LAYER ETE_TJ
  (* CLP SUBESTACAO (M262_Substacao) *)
  (* CLP LODO (M262_Lodo) *)
  (* CLP NEREDA (M262_Nereda) *)
  (* Painel Subestacao - Remota 1 (SUB_R1 .192), geradores QTAM1/QTAM2 (AGC150 .186/.187), MGE QGBT 220 V (.191) *)
  (* Agua de Reuso (1000) - Remota 2 (SUB_R2 .193), MGE .190 *)
  (* EEE Bruto (100) - Remota A1 (.197), inversores BS-100-01/02/03 (.200-.202), MGE .199 *)
  (* Pre-tratamento (200) - UCT_200_01 (.182), UCT_200_02 (.184), UCT_200_03 reserva; inversores BR-200-03/04 (.176/.177) *)
  (* Remota 2 do Nereda (NER_R2 .161, A12 canal 7) - lida pelo CLP Subestacao *)
  (* Gradeamento (100) - painel Vibropac (.207), comportas CO-100-01..04 (.203-.206) *)
  (* Sem painel definido - Dosagem de alcalinizante (800), sem campo *)
  (* Desinfeccao (700) - Remota A1, VC-700-01, UV Trojan, SC4500 pH/OD/turbidez, MGE .139 *)
  (* Lodo (900) - Remotas A2 (.135) e A10 (.136), inversores, valvulas e skids 900, MGE .246 *)
  (* Painel Nereda - Remotas A2/A10, Remota A11 (area do lodo: SludgeBuffer e Sludge Holding Tanks), sopradores Sulzer V4601-4604, SC1000/SC4500, inversores P4001-3/R4005/P4901-3, MGE .143 *)
  (* NEREDA REACTORS *)
  (* NEREDA PROCESS - HIDRYCO *)
  (* EMERGENCY RECIPIE *)
  (* NEREDA EQUIPMENT *)
  (* NEREDA AERATION *)
  (* INFLUENT FEED *)
  (* EFFLUENT *)
  (* SLUDGE BUFFER *)
  (* METAL SALT DOSING *)
  (* SLUDGE HOLDING TANK *)
  FBS
    EEEB : EEE_Bruto(cfgTempoFalhaBoiaL := 10, cfgTempoPartidaPressao := 30, cfgUsaFalhaComunicacao := TRUE, geradorConectado := TRUE); {SET_ATTRIBUTE(Configuration.Component.HideUnusedPorts, )}
    AGUA_REUSO : Agua_Reuso(cfgTempoBoia := 10, cfgBoiaInvertida := FALSE, cfgTempoCom := 5); {SET_ATTRIBUTE(Configuration.Component.HideUnusedPorts, )}
    SUBESTACAO : Subestacao(cfgTempoDiscordancia := 5, cfgTempoComGerador := 10, cfgTempoPulsoDisjuntor := 1, cfgTempoRespostaDisjuntor := 5); {SET_ATTRIBUTE(Configuration.Component.HideUnusedPorts, )}
    MGE_AGUA_REUSO : MGE_Generico(cfgTempoCom := 5); {SET_ATTRIBUTE(Configuration.Component.HideUnusedPorts, )}
    MGE_QGBT_220V : MGE_Generico(cfgTempoCom := 5); {SET_ATTRIBUTE(Configuration.Component.HideUnusedPorts, )}
    MGE_NEREDA : MGE_Generico(cfgTempoCom := 5); {SET_ATTRIBUTE(Configuration.Component.HideUnusedPorts, )}
    MGE_EEE_BRUTO : MGE_Generico(cfgTempoCom := 5); {SET_ATTRIBUTE(Configuration.Component.HideUnusedPorts, )}
    MGE_LODO : MGE_Generico(cfgTempoCom := 5); {SET_ATTRIBUTE(Configuration.Component.HideUnusedPorts, )}
    MGE_DESINFECCAO : MGE_Generico(cfgTempoCom := 5); {SET_ATTRIBUTE(Configuration.Component.HideUnusedPorts, )}
    Pre_Tratamento1 : UCT_PreTratamento(cfgInstalada := TRUE, cfgTempoCom := 10, cfgTempoReset := 2); {SET_ATTRIBUTE(Configuration.Component.HideUnusedPorts, )}
    Pre_Tratamento2 : UCT_PreTratamento(cfgInstalada := TRUE, cfgTempoCom := 10, cfgTempoReset := 2); {SET_ATTRIBUTE(Configuration.Component.HideUnusedPorts, )}
    Pre_Tratamento3 : UCT_PreTratamento(cfgInstalada := FALSE, cfgTempoCom := 10, cfgTempoReset := 2); {SET_ATTRIBUTE(Configuration.Component.HideUnusedPorts, )}
    FT_40_02 : Sensor_Generico(cfgUnidade := 'm3/h', cfgCasasDecimais := 1, cfgUsaConexao := TRUE, cfgComunicacao := FALSE, cfgNivel := FALSE, cfgBrutoMin := 4000.0, cfgBrutoMax := 20000.0, cfgFalhaMin := 3800.0, cfgFalhaMax := 22000.0, cfgTempoFalha := 5); {SET_ATTRIBUTE(Configuration.Component.HideUnusedPorts, )}
    DESINFECCAO : Desinfeccao_UV; {SET_ATTRIBUTE(Configuration.Component.HideUnusedPorts, )}
    DesidratacaoLodo : DesidratacaoLodo; {SET_ATTRIBUTE(Configuration.Component.HideUnusedPorts, )}
    EstocagemLodo : EstocagemLodo; {SET_ATTRIBUTE(Configuration.Component.HideUnusedPorts, )}
    Gradeamento : Gradeamento_Inovaisa; {SET_ATTRIBUTE(Configuration.Component.HideUnusedPorts, )}
    DosagemAlcalinizante : Dosagem_Alcalinizante; {SET_ATTRIBUTE(Configuration.Component.HideUnusedPorts, )}
    Mode : Mode; {SET_ATTRIBUTE(CompilerOptions, CheckConnectionsStrictly=False)}
    OpenWebPage : OpenWebPage(URL := 'http://192.168.1.10');
    OTHERS_DISCHARGE_VALVES_FB : OthersDischargeValves;
    EmergencyManagement : EmergencyManagement;
    Utilities : Utilities;
    EnergySignal : Frequency_Power;
    HeartBeat1 : HeartBeat;
    Aerator : NeredaCAeration;
    SludgeBuffer : NeredaSludgeBuffer_2;
    SludgeHoldingTank1 : SludgeHoldingTank;
    SludgeHoldingTank2 : SludgeHoldingTank;
    Reactor1 : NeredaReactor;
    Reactor2 : NeredaReactor;
    EmergencySB : EmergencySludgeBuffer;
    EmergencyReactor1 : EmergencyReactor_2;
    EmergencyReactor2 : EmergencyReactor_2;
    InfluentFeed : InfluentFeed;
  END_FBS
  EVENT_CONNECTIONS
    SUBESTACAO.921BB7D26016F39E TO EEEB.2B02D319AFE26590; (* planta nos geradores / bombas liberadas -> EEE Bruto *)
    SUBESTACAO.921BB7D26016F39E TO Pre_Tratamento1.0B595E2D755381E4;
    SUBESTACAO.921BB7D26016F39E TO Pre_Tratamento2.0B595E2D755381E4;
    SUBESTACAO.921BB7D26016F39E TO Pre_Tratamento3.0B595E2D755381E4;
    Pre_Tratamento1.5A6CC858EDC95420 TO Pre_Tratamento2.0B595E2D755381E4;
    Pre_Tratamento2.5A6CC858EDC95420 TO Pre_Tratamento3.0B595E2D755381E4;
    Pre_Tratamento3.5A6CC858EDC95420 TO EEEB.2B02D319AFE26590;
    EstocagemLodo.974B4969DB603762 TO DesidratacaoLodo.91E17855232378A8;
    EstocagemLodo.E3809710B35A5BE3 TO DesidratacaoLodo.335836E160C77742;
    DesidratacaoLodo.D64A39BCF02DDEB2 TO EstocagemLodo.AB5FAE61D1BCDDFE;
    DesidratacaoLodo.EA9A2427D178E8B5 TO EstocagemLodo.39F3DF7DDD7B4C23;
    DesidratacaoLodo.EE8958653A86D261 TO EstocagemLodo.4FA8CBCB1032FBD8;
    SUBESTACAO.921BB7D26016F39E TO DosagemAlcalinizante.3550FA6DB34A3727;
    SUBESTACAO.921BB7D26016F39E TO Gradeamento.D1B66AFAEC6D2FF0;
    SUBESTACAO.921BB7D26016F39E TO DESINFECCAO.3AA953731967D084;
    SUBESTACAO.921BB7D26016F39E TO Aerator.343299A527021480;
    SUBESTACAO.921BB7D26016F39E TO SludgeBuffer.9DD23EB33BCCE747;
    SUBESTACAO.921BB7D26016F39E TO InfluentFeed.9990B718E668E6B3;
    EstocagemLodo.3B317909428F66BD TO SludgeHoldingTank1.BD354E954D175C1F;
    EstocagemLodo.3B317909428F66BD TO SludgeHoldingTank2.BD354E954D175C1F;
    DosagemAlcalinizante.2549BCE0C5B3D328 TO Utilities.456D871DCB00F480;
  END_CONNECTIONS
  DATA_CONNECTIONS
    SUBESTACAO.FEF1963C61B73419 TO EEEB.D20C22571F86F121;
    SUBESTACAO.9CB30A27579CAC79 TO EEEB.B9262C2637F95B4A;
    SUBESTACAO.AD92EC25FAFA674A TO EEEB.011919C853DE622C;
    SUBESTACAO.F7B1C8F24F37DABA TO EEEB.EC0B0545A7F8DBEB;
    SUBESTACAO.5DB035BC4F7321F6 TO Pre_Tratamento1.D205F407BC981FB4;
    SUBESTACAO.FEF1963C61B73419 TO Pre_Tratamento1.2C19134423AEFFAA;
    SUBESTACAO.E3892FBEADB0545B TO Pre_Tratamento2.D205F407BC981FB4;
    SUBESTACAO.FEF1963C61B73419 TO Pre_Tratamento2.2C19134423AEFFAA;
    SUBESTACAO.85B535DFB1FB677D TO Pre_Tratamento3.D205F407BC981FB4;
    SUBESTACAO.FEF1963C61B73419 TO Pre_Tratamento3.2C19134423AEFFAA;
    Pre_Tratamento1.1F8CA54F12D8796B TO Pre_Tratamento2.3F3598C544A33E47;
    Pre_Tratamento1.A737D1113B918FC6 TO Pre_Tratamento2.BFB78C58CA08F906;
    Pre_Tratamento2.1F8CA54F12D8796B TO Pre_Tratamento3.3F3598C544A33E47;
    Pre_Tratamento2.A737D1113B918FC6 TO Pre_Tratamento3.BFB78C58CA08F906;
    Pre_Tratamento3.6948495C8744310C TO EEEB.83B944A122866558;
    EstocagemLodo.649314760363E488 TO DesidratacaoLodo.AC99B8EE5C6DBA64;
    EstocagemLodo.B87FCF9EF6E17A10 TO DesidratacaoLodo.D231A14376C3E2F6;
    EstocagemLodo.273D781A989DEA3F TO DesidratacaoLodo.DE00033B699DACF0;
    EstocagemLodo.0D2CE8145A8A40C5 TO DesidratacaoLodo.099E44A540EF9490;
    EstocagemLodo.E7A1F2C70FD2876B TO DesidratacaoLodo.426B37B9A495B79C;
    EstocagemLodo.5C0EE27FAC026E42 TO DesidratacaoLodo.FD17B98D889E4E9C;
    EstocagemLodo.28C5117F80A71252 TO DesidratacaoLodo.91FA512D1B0CCA17;
    EstocagemLodo.F39C9B782425030B TO DesidratacaoLodo.18A2A222BB911413;
    EstocagemLodo.CA5C991A51FB83CF TO DesidratacaoLodo.14561E73765FBECA;
    EstocagemLodo.5405EB7088EC4BDE TO DesidratacaoLodo.1CD77F0C67EACF01;
    DesidratacaoLodo.317BB96205F3F911 TO EstocagemLodo.EE49B187C469C0B7;
    DesidratacaoLodo.A2D8149F0FE69321 TO EstocagemLodo.E59CBDC75C3131D4;
    DesidratacaoLodo.08464482A0BF6120 TO EstocagemLodo.8E87331950BD000E;
    DesidratacaoLodo.4080C84A5DF2BAE8 TO EstocagemLodo.3B31F82669E06299;
    SUBESTACAO.B9F74BEEB26000F4 TO DosagemAlcalinizante.A0398C4E77A10EEE;
    SUBESTACAO.499BDAC4EA9F62DF TO DosagemAlcalinizante.7CA01E1D24150792;
    SUBESTACAO.FEF1963C61B73419 TO DosagemAlcalinizante.7838A99D6B60D295;
    SUBESTACAO.2BBFC35BA4EC9BC5 TO Gradeamento.358F3774D14189DB;
    SUBESTACAO.FEF1963C61B73419 TO Gradeamento.98A20843E1C25CF2;
    SUBESTACAO.45C7CD3C2C5255A5 TO DESINFECCAO.B6FA6DECDD9ED22F;
    SUBESTACAO.A0BFF3F0BE735315 TO DESINFECCAO.FE5067C199042FFC;
    SUBESTACAO.FEF1963C61B73419 TO DESINFECCAO.29FAEE93999A7375;
    DesidratacaoLodo.9DCD88E1901DA328 TO EstocagemLodo.A8767255ECC4E3FD;
    SUBESTACAO.28CCDBC73D782726 TO Aerator.E8E5FF489B43618A;
    SUBESTACAO.5F05D9810446E7DA TO Aerator.A6249B75BAECD359;
    SUBESTACAO.62B1CE99737B56B7 TO Aerator.9706F98C2A856240;
    SUBESTACAO.D53B21982E1C7690 TO Aerator.639EFA592CF3B7AB;
    SUBESTACAO.FEF1963C61B73419 TO Aerator.B6004AB02CFE077D;
    SUBESTACAO.38835B908E410028 TO SludgeBuffer.7D03DBDF71B8C2FE;
    SUBESTACAO.60DD75A9AF1A4BF6 TO SludgeBuffer.D58F38BFC1670450;
    SUBESTACAO.5A0597290C490F4A TO SludgeBuffer.5CEDBAD4251CEB62;
    SUBESTACAO.FEF1963C61B73419 TO SludgeBuffer.169E5A2DB0450A6B;
    SUBESTACAO.B81B83BF98ACFA31 TO InfluentFeed.FB134FF10099DEF1;
    SUBESTACAO.BD12E9799143BEA9 TO InfluentFeed.2D5BC448F9BDE10B;
    SUBESTACAO.FEF1963C61B73419 TO InfluentFeed.4BFFE021F8C35676;
    EstocagemLodo.E2CA55FAEBB4E606 TO SludgeHoldingTank1.875A0A21AD0E0927;
    EstocagemLodo.5FECFF6590BA1CB8 TO SludgeHoldingTank1.51A296D74729C981;
    EstocagemLodo.C03F8F23B8219B89 TO SludgeHoldingTank1.88E72593FBD99CC6;
    EstocagemLodo.47DA0D3EDA2667D7 TO SludgeHoldingTank2.875A0A21AD0E0927;
    EstocagemLodo.5EDEC437D5610CDE TO SludgeHoldingTank2.51A296D74729C981;
    EstocagemLodo.D43E44FA212AEC2C TO SludgeHoldingTank2.88E72593FBD99CC6;
    DosagemAlcalinizante.102C84667EC49B91 TO Utilities.380D19E58AADF575;
    DosagemAlcalinizante.32CD2F3F12A90B15 TO Utilities.B240C89A22FE0002;
  END_CONNECTIONS
  ADAPTER_CONNECTIONS
    HeartBeat1.40 TO Mode.6E012D59F948069E;
    Mode.50 TO SludgeBuffer.6D7943A09F73313C;
    Reactor1.0FAC572B8C8842D9 TO EmergencyReactor1.850ED619A957D063;
    Reactor2.0FAC572B8C8842D9 TO EmergencyReactor2.850ED619A957D063;
    InfluentFeed.06B5BF90025137D8 TO SludgeBuffer.04BD059D1BCDA8FF;
    InfluentFeed.08DA021DBE2FF670 TO SludgeBuffer.34E82C716D68805B;
    SludgeHoldingTank1.745E7C7F86CD93D6 TO SludgeBuffer.1369AAF8C65D025F;
    SludgeHoldingTank2.745E7C7F86CD93D6 TO SludgeBuffer.103390B72A3B733A;
    OTHERS_DISCHARGE_VALVES_FB.82A979F8A1C1CE4A TO Reactor1.AE9DB11716461BE5;
    OTHERS_DISCHARGE_VALVES_FB.00DDB30B96836B1C TO Reactor2.AE9DB11716461BE5;
    Mode.39 TO Reactor1.8E8BC8CAE0ABBEF0;
    Mode.40 TO Reactor2.8E8BC8CAE0ABBEF0;
    Mode.55 TO EmergencyManagement.FA37C5C7FF880AB4;
    Reactor1.53509993DCC2E69E TO EmergencyManagement.03E1DF24854B5087;
    Reactor2.53509993DCC2E69E TO EmergencyManagement.8D40980BCD10D06B;
    EmergencyManagement.5C1263F1F6F0F578 TO EmergencyReactor1.73503C83163B2D86;
    EmergencyManagement.6B6FC4EBFE551754 TO EmergencyReactor2.73503C83163B2D86;
    Reactor1.E962C7AC1C669349 TO Aerator.IBlowerReactor;
    Reactor2.E962C7AC1C669349 TO Aerator.036B0699AE92B07E;
    Reactor1.EF12C2F0857E0401 TO InfluentFeed.458126F8619187E9;
    Reactor2.EF12C2F0857E0401 TO InfluentFeed.13A00CB3B1B3C5BD;
    EmergencyReactor1.ADE9AC252194767E TO Reactor1.4FE3E9A63522A043;
    EmergencyReactor2.ADE9AC252194767E TO Reactor2.4FE3E9A63522A043;
    SludgeBuffer.5220CD4AB4D5EF57 TO Reactor1.64A5E847CFF537B2;
    SludgeBuffer.F8A56E33E99EA0E4 TO Reactor2.64A5E847CFF537B2;
    SludgeBuffer.2EF6B69B645AE6E1 TO InfluentFeed.9135BA3E72B25810;
    EmergencyManagement.10001B393681040B TO OTHERS_DISCHARGE_VALVES_FB.0FC638121CDA6752;
    SludgeBuffer.8B97DDD2DF3E853F TO EmergencyManagement.92B17EFA7CB0DA14;
    EmergencyReactor2.D6CF55AACA664FB9 TO EmergencySB.A9597B321AC24B8F;
    EmergencyReactor1.D6CF55AACA664FB9 TO EmergencySB.E201588BE0264C59;
    InfluentFeed.072EC58E32F5B902 TO Reactor1.9D6CC0A1E886795A;
    InfluentFeed.57887779F0B6E332 TO Reactor2.9D6CC0A1E886795A;
    SludgeBuffer.0CE6DD66A1C58D5B TO Reactor1.6D054A47338EC161;
    SludgeBuffer.DE069E6752438E1A TO Reactor2.6D054A47338EC161;
    EmergencySB.CC52284A3E90E837 TO SludgeBuffer.8642DEF89CD05FB2;
    InfluentFeed.091DBEAA531EFD46 TO EmergencyManagement.547ED878E258385C;
  END_CONNECTIONS
END_LAYER
